// TIA Portal V21 export
DATA_BLOCK "F_IDB_MainSafety"   // DB2, F_DB
NAME : FUSI
// stored: InstanceOfName F_FB_MainSafety, InstanceOfType FB
"F_FB_MainSafety"
   // VAR
   //    Enable : Bool;
   //    Released : Bool;
   //    LogicRelease : Bool;
   // END_VAR
BEGIN
END_DATA_BLOCK
